Fanuc KAREL source: KT00155.KL

PROGRAM KT00155
%NOLOCKGROUP
VAR
  H1: ARRAY[2] OF SHORT
  R2: REAL
  OUT: INTEGER
BEGIN
  H1[1] = 2
    R2 = 3.0
  OUT = H1[1] DIV R2
END KT00155
